{region 'Documentation'}
(*!
<summary>Checks equality with the expected TIME value.</summary>
*)
{endregion}
FUNCTION_BLOCK AssertEqual_Time EXTENDS AssertionBase
VAR_INPUT
    IN : TIME; //! Actual value checked or observed by this Assertion.
    Expected : TIME; //! Reference value for comparison with IN.
END_VAR

SUPER^();

{region 'Documentation'}
(*!
<summary>Evaluate the typed duration relation and report higher-priority errors first.</summary>
*)
{endregion}
METHOD PROTECTED Assert
VAR
    Message : STRING(GVL_Constants.MessageLength);
    ExpectedText : STRING(GVL_Constants.AssertionValueLength);
    ActualText : STRING(GVL_Constants.AssertionValueLength);
END_VAR
IF NOT EvaluationActive THEN
    RETURN;
END_IF;

IF Result = E_Result.Error THEN
    RETURN;
END_IF;

IF Result = E_Result.Failed THEN
    RETURN;
END_IF;

IF IN <> Expected THEN
    ExpectedText := TIME_TO_STRING(Expected);
    ActualText := TIME_TO_STRING(IN);
    Message := CONCAT('Assertion failed: values are not equal. Expected = ',
        ExpectedText);
    Message := CONCAT(Message, ', Actual = ');
    Message := CONCAT(Message, ActualText);
    Message := CONCAT(Message, '.');
    Fail(Message := Message);
    RETURN;
END_IF;

Pass();
END_METHOD

END_FUNCTION_BLOCK

(* stored: Version 1.1.0.1
   POU AssertEqual_Time: Id {1f1b2c09-418c-4977-b7a7-1604df8794ce}, SpecialFunc None
   Folder Internal: Id {0035f1e8-8fea-4c65-8d6c-ca142b9e89e3}
   Method Assert: Id {f01ca648-7e0e-481c-8dd7-55fd88739990} *)
